// TIA Portal V21 export
// export: Created 2026-11-10T19:21:33.8745756Z, ExportSetting WithDefaults, DisplayName Totally Integrated Automation Portal, DisplayVersion V21 Update 3, DisplayName STEP 7 Professional, DisplayVersion V21 Update 3, DisplayName STEP 7 Safety, DisplayVersion V21, DisplayName Tech WebApplication, DisplayVersion V21, DisplayName WinCC Basic/Comfort/Advanced, DisplayVersion V21 Update 3, DisplayName WinCC Unified, DisplayVersion V21 Update 3
FUNCTION_BLOCK "FB_Lad_us004"   // FB4, LAD
{ S7_Optimized_Access := 'TRUE' }
VERSION : 0.1
// stored: AutoNumber true, IsIECCheckEnabled false, IsRetainMemResEnabled false, MemoryReserve 100, SetENOAutomatically false, UDAEnableTagReadback false
   VAR_INPUT
      v_run : Bool;
      v_off2 : Bool;
      v_off3 : Bool;
      v_f_ack : Bool;
      v_dir : Bool;
      v_drive : USInt;
      v_pzd_len : USInt;
      v_speed_sp : Real;
      v_ctrl3 : Word;
      v_ctrl4 : Word;
      v_ctrl5 : Word;
      v_ctrl6 : Word;
      v_ctrl7 : Word;
      v_ctrl8 : Word;
   END_VAR
   VAR_OUTPUT
      v_ndr : Bool;
      v_error : Bool;
      v_status : Word;
      v_run_en : Bool;
      v_d_dir : Bool;
      v_inhibit : Bool;
      v_fault : Bool;
      v_speed : Real;
      v_status1 : Word;
      v_status3 : Word;
      v_status4 : Word;
      v_status5 : Word;
      v_status6 : Word;
      v_status7 : Word;
      v_status8 : Word;
   END_VAR
   VAR
      inst { S7_SetPoint := 'True'} : USS_Drive_Control;
   END_VAR
BEGIN

REGION Network 1: USS_DRIVE - Swap data with drive
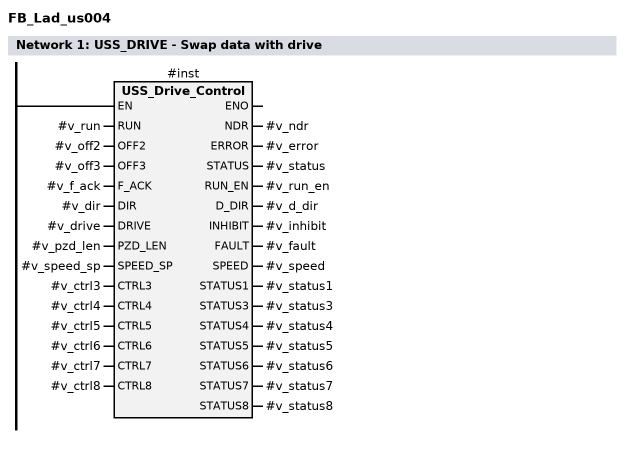
   RUNG wire#powerrail
      #inst.USS_Drive_Control(RUN := #v_run, OFF2 := #v_off2, OFF3 := #v_off3, F_ACK := #v_f_ack, DIR := #v_dir, DRIVE := #v_drive, PZD_LEN := #v_pzd_len, SPEED_SP := #v_speed_sp, CTRL3 := #v_ctrl3, CTRL4 := #v_ctrl4, CTRL5 := #v_ctrl5, CTRL6 := #v_ctrl6, CTRL7 := #v_ctrl7, CTRL8 := #v_ctrl8, NDR => #v_ndr, ERROR => #v_error, STATUS => #v_status, RUN_EN => #v_run_en, D_DIR => #v_d_dir, INHIBIT => #v_inhibit, FAULT => #v_fault, SPEED => #v_speed, STATUS1 => #v_status1, STATUS3 => #v_status3, STATUS4 => #v_status4, STATUS5 => #v_status5, STATUS6 => #v_status6, STATUS7 => #v_status7, STATUS8 => #v_status8)
   END_RUNG
   // the same network as SCL:
   #inst(RUN := #v_run,   // USS_Drive_Control
         OFF2 := #v_off2,
         OFF3 := #v_off3,
         F_ACK := #v_f_ack,
         DIR := #v_dir,
         DRIVE := #v_drive,
         PZD_LEN := #v_pzd_len,
         SPEED_SP := #v_speed_sp,
         CTRL3 := #v_ctrl3,
         CTRL4 := #v_ctrl4,
         CTRL5 := #v_ctrl5,
         CTRL6 := #v_ctrl6,
         CTRL7 := #v_ctrl7,
         CTRL8 := #v_ctrl8,
         NDR => #v_ndr,
         ERROR => #v_error,
         STATUS => #v_status,
         RUN_EN => #v_run_en,
         D_DIR => #v_d_dir,
         INHIBIT => #v_inhibit,
         FAULT => #v_fault,
         SPEED => #v_speed,
         STATUS1 => #v_status1,
         STATUS3 => #v_status3,
         STATUS4 => #v_status4,
         STATUS5 => #v_status5,
         STATUS6 => #v_status6,
         STATUS7 => #v_status7,
         STATUS8 => #v_status8);
END_REGION
END_FUNCTION_BLOCK
